(* IEC 61131-3 sources: BODAS-HelloWorld/st/bodas_rc18_12_40/plc_logic/application/01_maintask/10_service/programs, 5 files *)

(* ---- uds_diag_chklvl-UDS_Diag_ChkLvl.st ---- *)
(* --- Interface --- *)
(*********************************************************************************************************************
 *     __   __   ___  ___           __   __        __   __  ___
 *   /_ / /  / /__  /    /__/     /_ / /_   |_ / /_ / /  /  /  /__/
 *  /__/ /__/ __ / /__  /  /     /  | /__  /  | /  | /__/  /  /  /
 *
 * Project: Hello World for ml290.rts
 *
 * Function: UDS_Diag_ChkLvl
 *
 * Author:
 *
 * Description:
 * Function for level check
 *
 * (c) Copyright by BOSCH REXROTH AG, all rights reserved
 *
 *********************************************************************************************************************)
FUNCTION UDS_Diag_ChkLvl : USINT
VAR_INPUT
	i_Mask_u32  : UDINT;
	i_Level_u16 : UINT;
END_VAR

(* --- Implementation --- *)
(*UDS_Diag_ChkLvl := GVL_UDS.UDS_NEGATIVE_RESPONSE;*)
UDS_Diag_ChkLvl := 1;

(* First check security as defined in ISO 14229 - see bds_sec_accessLevel_te *)
IF (0 <> (UDINT_TO_WORD(i_Mask_u32) AND SHL(i_Level_u16, 16#1))) THEN
	(*UDS_Diag_ChkLvl := GVL_UDS.UDS_POSITIVE_RESPONSE;*)
	UDS_Diag_ChkLvl := 0;
ELSE
	;
END_IF

(* ---- uds_readcallback-UDS_ReadCallback.st ---- *)
(* --- Interface --- *)
FUNCTION UDS_ReadCallback
VAR_INPUT
	//a variable to which the content has to be written
	UDSReadData_pau8 : POINTER TO USINT;
END_VAR
VAR
	// variables for internal operations
	//data_au8 : ARRAY[0..8] OF BYTE;
	i                     : BYTE;
	DidValue_u16          : UINT;
	set_u8                : USINT;
	ret_secLevel          : UINT;
	Level_pu16            : POINTER TO UINT;
	ret_response          : BOOL;
	temp_sec_level        : BOOL;
	uPmpSnsr_mV_u16       : UINT;
	fctPmp_s16            : INT;
	stBrkSwt_u8           : USINT;
	iPmpFwdAct_mA_u16     : UINT;
	funcRet_u8            : USINT;
	UDSReadData_pau8_poby : POINTER TO ARRAY[0..7] OF BYTE;
	UDSReadData_pau8_by   : ARRAY[0..7] OF BYTE;
	DID_0103_s32          : DINT;
	DiagChkLvlRet_u8      : USINT;
END_VAR

(* --- Implementation --- *)
(* Get the DID requested by tester present *)
bds_uds_GetActiveDid(ADR(DidValue_u16));

//bds_can_sendData(bds_can_Chnl_te.BDS_CAN_1_D, 5, BDS_CAN_EXD_DU8, 2, ADR(DidValue_u16));
//CASE DidValue_u16 OF
// 16#C003, 16#D001, 16#D002:
(* here check th security level *)
//bds_sec_getLevel(BDS_SEC_ASW_INST_NAME_2_E, ADR(Level_pu16));
//DiagChkLvlRet_u8 := UDS_Diag_ChkLvl(16#00000004, Level_pu16^);
//ELSE
(* all levels allowed *)
//bds_sec_getLevel(BDS_SEC_ASW_INST_NAME_1_E, ADR(Level_pu16));
//DiagChkLvlRet_u8 := UDS_Diag_ChkLvl(16#FFFFFFFF, Level_pu16^);
//DiagChkLvlRet_u8 := 0;
//END_CASE
IF (TRUE) THEN
	//IF( NOT( USINT_TO_BOOL( DiagChkLvlRet_u8 ) ) ) THEN
	CASE DidValue_u16 OF
	(* Handle the read operation at DIDs *)
	(* Parameters *)
	16#C001: bds_uds_setCallbackStatus(0); (* E_OK *)
		UDSReadData_pau8[1] := INT_TO_BYTE(SHR(GlobalVariables.PrmAsw_gstruc.fctPmp_s16, 8));
		UDSReadData_pau8[0] := INT_TO_BYTE(GlobalVariables.PrmAsw_gstruc.fctPmp_s16);
	16#C002: bds_uds_setCallbackStatus(0); (* E_OK *)
		UDSReadData_pau8[1] := TO_BYTE(SHR(GlobalVariables.PrmAsw_gstruc.listCtrlVlv_enu, 8));
		UDSReadData_pau8[0] := TO_BYTE(GlobalVariables.PrmAsw_gstruc.listCtrlVlv_enu);
	16#C003: bds_uds_setCallbackStatus(0); (* E_OK *)
		UDSReadData_pau8[1] := INT_TO_BYTE(SHR(GlobalVariables.PrmAsw_gstruc.nrCogs_s16, 8));
		UDSReadData_pau8[0] := INT_TO_BYTE(GlobalVariables.PrmAsw_gstruc.nrCogs_s16);
	16#01C7: bds_uds_setCallbackStatus(0); (* E_OK *)
		UDSReadData_pau8[1] := UINT_TO_BYTE(SHR(GlobalVariables.PrmAsw_gstruc.iSpSafout1_u16, 8));
		UDSReadData_pau8[0] := UINT_TO_BYTE(GlobalVariables.PrmAsw_gstruc.iSpSafout1_u16);
	16#01C8: bds_uds_setCallbackStatus(0); (* E_OK *)
		UDSReadData_pau8[1] := UINT_TO_BYTE(SHR(GlobalVariables.PrmAsw_gstruc.iSpSafout2_u16, 8));
		UDSReadData_pau8[0] := UINT_TO_BYTE(GlobalVariables.PrmAsw_gstruc.iSpSafout2_u16);
	16#D001: bds_uds_setCallbackStatus(0); (* E_OK *)
		UDSReadData_pau8[0] := BOOL_TO_BYTE(GlobalVariables.PrmAsw_gstruc.PrmDbg_struc.flgXcpOn_b);
	16#D002: bds_uds_setCallbackStatus(0); (* E_OK *)
		UDSReadData_pau8[0] := BOOL_TO_BYTE(GlobalVariables.PrmAsw_gstruc.PrmDbg_struc.flgStoreDataToNvm_b);
	16#C010: bds_uds_setCallbackStatus(0); (* E_OK *)
		UDSReadData_pau8[1] := UINT_TO_BYTE(SHR(GlobalVariables.PrmAsw_gstruc.eff_perc_au16[0], 8));
		UDSReadData_pau8[0] := UINT_TO_BYTE(GlobalVariables.PrmAsw_gstruc.eff_perc_au16[0]);
		UDSReadData_pau8[3] := UINT_TO_BYTE(SHR(GlobalVariables.PrmAsw_gstruc.eff_perc_au16[1], 8));
		UDSReadData_pau8[2] := UINT_TO_BYTE(GlobalVariables.PrmAsw_gstruc.eff_perc_au16[1]);
		UDSReadData_pau8[5] := UINT_TO_BYTE(SHR(GlobalVariables.PrmAsw_gstruc.eff_perc_au16[2], 8));
		UDSReadData_pau8[4] := UINT_TO_BYTE(GlobalVariables.PrmAsw_gstruc.eff_perc_au16[2]);
	16#C020: bds_uds_setCallbackStatus(0); (* E_OK *)
		UDSReadData_pau8[1] := UINT_TO_BYTE(SHR(GlobalVariables.PrmAsw_gstruc.nEngSpd_rpm_au16[0], 8));
		UDSReadData_pau8[0] := UINT_TO_BYTE(GlobalVariables.PrmAsw_gstruc.nEngSpd_rpm_au16[0]);
		UDSReadData_pau8[3] := UINT_TO_BYTE(SHR(GlobalVariables.PrmAsw_gstruc.nEngSpd_rpm_au16[1], 8));
		UDSReadData_pau8[2] := UINT_TO_BYTE(GlobalVariables.PrmAsw_gstruc.nEngSpd_rpm_au16[1]);
		UDSReadData_pau8[5] := UINT_TO_BYTE(SHR(GlobalVariables.PrmAsw_gstruc.nEngSpd_rpm_au16[2], 8));
		UDSReadData_pau8[4] := UINT_TO_BYTE(GlobalVariables.PrmAsw_gstruc.nEngSpd_rpm_au16[2]);
	(* Process Values *)
	16#A001: bds_uds_setCallbackStatus(0); (* E_OK *)
		UDSReadData_pau8[1] := UINT_TO_BYTE(SHR(PRG_Inputs.uPmpSnsr_mV_u16, 8));
		UDSReadData_pau8[0] := UINT_TO_BYTE(PRG_Inputs.uPmpSnsr_mV_u16);
	16#A002: bds_uds_setCallbackStatus(0); (* E_OK *)
		UDSReadData_pau8[0] := INT_TO_BYTE(PRG_Outputs.st_BrkSwt_u8);
	16#A003: bds_uds_setCallbackStatus(0); (* E_OK *)
		UDSReadData_pau8[1] := UDINT_TO_BYTE(SHR(PRG_Inputs.frqVehSnsr_Hz_u32, 8));
		UDSReadData_pau8[0] := UDINT_TO_BYTE(PRG_Inputs.frqVehSnsr_Hz_u32);
	16#B001: bds_uds_setCallbackStatus(0); (* E_OK *)
		UDSReadData_pau8[1] := UINT_TO_BYTE(SHR(PRG_Outputs.no_CurrentK07_mA_u16, 8));
		UDSReadData_pau8[0] := UINT_TO_BYTE(PRG_Outputs.no_CurrentK07_mA_u16);
	16#B002: bds_uds_setCallbackStatus(0); (* E_OK *)
		UDSReadData_pau8[0] := PRG_Outputs.st_CtrlValve_u8;
	16#B003: bds_uds_setCallbackStatus(0); (* E_OK *)
		UDSReadData_pau8[1] := UINT_TO_BYTE(SHR(PRG_Inputs.vWhlSpd_kph_u16, 8));
		UDSReadData_pau8[0] := UINT_TO_BYTE(PRG_Inputs.vWhlSpd_kph_u16);
		ELSE
			bds_uds_setCallbackStatus(1); (* E_OK *)
	END_CASE
ELSE
	bds_uds_setCallbackStatus(1); (* E_NOK *)
END_IF

(* ---- uds_writecallback-UDS_WriteCallback.st ---- *)
(* --- Interface --- *)
FUNCTION UDS_WriteCallback
VAR_INPUT
	UDSReadData_pau8 : POINTER TO USINT;
END_VAR
VAR
	DidValue_u16     : UINT;
	DiagChkLvlRet_u8 : USINT;
	Level_pu8        : POINTER TO USINT;
END_VAR

(* --- Implementation --- *)
(* Get the DID requested by tester present *)
bds_uds_GetActiveDid(ADR(DidValue_u16));

(* here check the security level *)
CASE DidValue_u16 OF
16#C003, 16#D001, 16#D002:
	(* security level 2 *)
	//bds_sec_getLevel(BDS_SEC_ASW_INST_NAME_1_E, ADR(Level_pu8));
	//DiagChkLvlRet_u8 := UDS_Diag_ChkLvl(16#00000004, Level_pu8^);
	DiagChkLvlRet_u8 := 0;
	ELSE
		(*bds_sec_getLevel(BDS_SEC_ASW_INST_NAME_1_E, ADR(Level_pu8));
	DiagChkLvlRet_u8 := UDS_Diag_ChkLvl(16#FFFFFFFF, Level_pu8^);*)
		DiagChkLvlRet_u8 := 0;
END_CASE

IF (NOT (USINT_TO_BOOL(DiagChkLvlRet_u8))) THEN
	CASE DidValue_u16 OF
	(* Handle the write operation at DID 0xC001 *)
	16#C001: bds_uds_setCallbackStatus(0); (* E_OK *)
		GlobalVariables.PrmAsw_gstruc.fctPmp_s16 := WORD_TO_INT(USINT_TO_WORD(UDSReadData_pau8[0]) + SHL(USINT_TO_WORD(UDSReadData_pau8[1]), 8));
	(* Handle the write operation at DID 0xC002 *)
	16#C002: bds_uds_setCallbackStatus(0); (* E_OK *)
		GlobalVariables.PrmAsw_gstruc.listCtrlVlv_enu.0 := UDSReadData_pau8[0].0;
		GlobalVariables.PrmAsw_gstruc.listCtrlVlv_enu.1 := UDSReadData_pau8[0].1;
		GlobalVariables.PrmAsw_gstruc.listCtrlVlv_enu.2 := UDSReadData_pau8[0].2;
		GlobalVariables.PrmAsw_gstruc.listCtrlVlv_enu.3 := UDSReadData_pau8[0].3;
		GlobalVariables.PrmAsw_gstruc.listCtrlVlv_enu.4 := UDSReadData_pau8[0].4;
		GlobalVariables.PrmAsw_gstruc.listCtrlVlv_enu.5 := UDSReadData_pau8[0].5;
		GlobalVariables.PrmAsw_gstruc.listCtrlVlv_enu.6 := UDSReadData_pau8[0].6;
		GlobalVariables.PrmAsw_gstruc.listCtrlVlv_enu.7 := UDSReadData_pau8[0].7;
	(* Handle the write operation at DID 0xC003 *)
	16#C003: bds_uds_setCallbackStatus(0); (* E_OK *)
		GlobalVariables.PrmAsw_gstruc.nrCogs_s16 := WORD_TO_INT(USINT_TO_WORD(UDSReadData_pau8[0]) + SHL(USINT_TO_WORD(UDSReadData_pau8[1]), 8));
	(* Handle the write operation at DID 0x01C7 *)
	16#01C7: bds_uds_setCallbackStatus(0); (* E_OK *)
		GlobalVariables.PrmAsw_gstruc.iSpSafout1_u16 :=
			WORD_TO_UINT(USINT_TO_WORD(UDSReadData_pau8[0]) + SHL(USINT_TO_WORD(UDSReadData_pau8[1]), 8));
	(* Handle the write operation at DID 0x01C8 *)
	16#01C8: bds_uds_setCallbackStatus(0); (* E_OK *)
		GlobalVariables.PrmAsw_gstruc.iSpSafout2_u16 :=
			WORD_TO_UINT(USINT_TO_WORD(UDSReadData_pau8[0]) + SHL(USINT_TO_WORD(UDSReadData_pau8[1]), 8));
	(* Handle the write operation at DID 0xD001 *)
	16#D001: bds_uds_setCallbackStatus(0); (* E_OK *)
		GlobalVariables.PrmAsw_gstruc.PrmDbg_struc.flgXcpOn_b := USINT_TO_BOOL(UDSReadData_pau8[0]);
	(* Handle the write operation at DID 0xD002 *)
	16#D002: bds_uds_setCallbackStatus(0); (* E_OK *)
		GlobalVariables.PrmAsw_gstruc.PrmDbg_struc.flgStoreDataToNvm_b := USINT_TO_BOOL(UDSReadData_pau8[0]);
	(* Handle the write operation at DID 0xC010 *)
	16#C010: bds_uds_setCallbackStatus(0); (* E_OK *)
		//GlobalVariables.PrmAsw_gstruc.eff_perc_au16[0] := WORD_TO_UINT(USINT_TO_WORD(UDSReadData_pau8[0]) + SHL(USINT_TO_WORD(UDSReadData_pau8[1]), 8));
		//GlobalVariables.PrmAsw_gstruc.eff_perc_au16[1] := WORD_TO_UINT(USINT_TO_WORD(UDSReadData_pau8[2]) + SHL(USINT_TO_WORD(UDSReadData_pau8[3]), 8));
		//GlobalVariables.PrmAsw_gstruc.eff_perc_au16[2] := WORD_TO_UINT(USINT_TO_WORD(UDSReadData_pau8[4]) + SHL(USINT_TO_WORD(UDSReadData_pau8[5]), 8));
	(* Handle the write operation at DID 0xC020 *)
	16#C020:
			//GlobalVariables.PrmAsw_gstruc.nEngSpd_rpm_au16[0] := WORD_TO_UINT(USINT_TO_WORD(UDSReadData_pau8[0]) + SHL(USINT_TO_WORD(UDSReadData_pau8[1]), 8));
			//GlobalVariables.PrmAsw_gstruc.nEngSpd_rpm_au16[1] := WORD_TO_UINT(USINT_TO_WORD(UDSReadData_pau8[2]) + SHL(USINT_TO_WORD(UDSReadData_pau8[3]), 8));
			//GlobalVariables.PrmAsw_gstruc.nEngSpd_rpm_au16[2] := WORD_TO_UINT(USINT_TO_WORD(UDSReadData_pau8[4]) + SHL(USINT_TO_WORD(UDSReadData_pau8[5]), 8));
		ELSE
			bds_uds_setCallbackStatus(1); (* E_NOK *)
	END_CASE
ELSE
	bds_uds_setCallbackStatus(1); (* E_NOK *)
END_IF

(* ---- uds_defaultcallback-UDS_DefaultCallback.st ---- *)
(* --- Interface --- *)
PROGRAM UDS_DefaultCallback
VAR
END_VAR

(* --- Implementation --- *)
GlobalVariables.PrmAsw_gstruc.fctPmp_s16                       := GlobalVariables.PrmAsw_cgstruc.fctPmp_s16;
GlobalVariables.PrmAsw_gstruc.listCtrlVlv_enu                  := GlobalVariables.PrmAsw_cgstruc.listCtrlVlv_enu;
GlobalVariables.PrmAsw_gstruc.nrCogs_s16                       := GlobalVariables.PrmAsw_cgstruc.nrCogs_s16;
GlobalVariables.PrmAsw_gstruc.iSpSafout1_u16                   := GlobalVariables.PrmAsw_cgstruc.iSpSafout1_u16;
GlobalVariables.PrmAsw_gstruc.iSpSafout2_u16                   := GlobalVariables.PrmAsw_cgstruc.iSpSafout2_u16;
GlobalVariables.PrmAsw_gstruc.PrmDbg_struc.flgXcpOn_b          := GlobalVariables.PrmAsw_cgstruc.PrmDbg_struc.flgXcpOn_b;
GlobalVariables.PrmAsw_gstruc.PrmDbg_struc.flgStoreDataToNvm_b := GlobalVariables.PrmAsw_cgstruc.PrmDbg_struc.flgStoreDataToNvm_b;
GlobalVariables.PrmAsw_gstruc.eff_perc_au16[0]                 := GlobalVariables.PrmAsw_cgstruc.eff_perc_au16[0];
GlobalVariables.PrmAsw_gstruc.eff_perc_au16[1]                 := GlobalVariables.PrmAsw_cgstruc.eff_perc_au16[1];
GlobalVariables.PrmAsw_gstruc.eff_perc_au16[2]                 := GlobalVariables.PrmAsw_cgstruc.eff_perc_au16[2];
GlobalVariables.PrmAsw_gstruc.nEngSpd_rpm_au16[0]              := GlobalVariables.PrmAsw_cgstruc.nEngSpd_rpm_au16[0];
GlobalVariables.PrmAsw_gstruc.nEngSpd_rpm_au16[1]              := GlobalVariables.PrmAsw_cgstruc.nEngSpd_rpm_au16[1];
GlobalVariables.PrmAsw_gstruc.nEngSpd_rpm_au16[2]              := GlobalVariables.PrmAsw_cgstruc.nEngSpd_rpm_au16[2];

(* ---- uds_routinecallback-UDS_RoutineCallback.st ---- *)
(* --- Interface --- *)
PROGRAM UDS_RoutineCallback
VAR
	NvmWriteRet_u16  : UINT;
	DiagChkLvlRet_u8 : USINT;
	Level_pu8        : POINTER TO USINT;
END_VAR

(* --- Implementation --- *)
(* here check th security level *)
//bds_sec_getLevel(BDS_SEC_ASW_INST_NAME_1_E, ADR(Level_pu8));
//DiagChkLvlRet_u8 := UDS_Diag_ChkLvl(16#00000004, Level_pu8^);
DiagChkLvlRet_u8 := 0;

IF (NOT (USINT_TO_BOOL(DiagChkLvlRet_u8))) THEN
	NvmWriteRet_u16 :=
		bds_mem_writeBlock(UINT_TO_USINT(bds_mem_nvmBlock01_512_R_D), ADR(GlobalVariables.PrmAsw_gstruc), 0, SIZEOF(GlobalVariables.PrmAsw_gstruc));

	IF (0 = NvmWriteRet_u16) THEN
		bds_uds_setCallbackStatus(0); (* E_OK *)
	ELSE
		bds_uds_setCallbackStatus(10); (* E_NOK which decrements to 1. i.e executes for 10 cycles before E_NOK is set ( wait time ill date is written to NVM) *)
	END_IF
ELSE
	bds_uds_setCallbackStatus(10); (* E_NOK *)
END_IF
